PROGRAM main
  VAR
    B1 AT %IX0.0   : BOOL; (* sensor de cajas *)
    KM1 AT %QX0.0  : BOOL; (* banda (bobina 00001 para la PC) *)
    CAJAS AT %MW0  : INT; (* holding 40001: cajas contadas *)
    MARCHA AT %MW1 : INT; (* holding 40002: marcha, la escribe la PC *)
    META AT %MW2   : INT; (* holding 40003: meta de cajas, la escribe la PC *)
    F_CAJA         : R_TRIG;
    CAJA           : BOOL; (* flanco de B1 *)
  END_VAR
  VAR  (* added by the conversion: wires and edge detectors of the diagram *)
    _ADD7_OUT : INT;
    _SEL4_OUT : INT;
    _NE11_OUT : BOOL;
  END_VAR

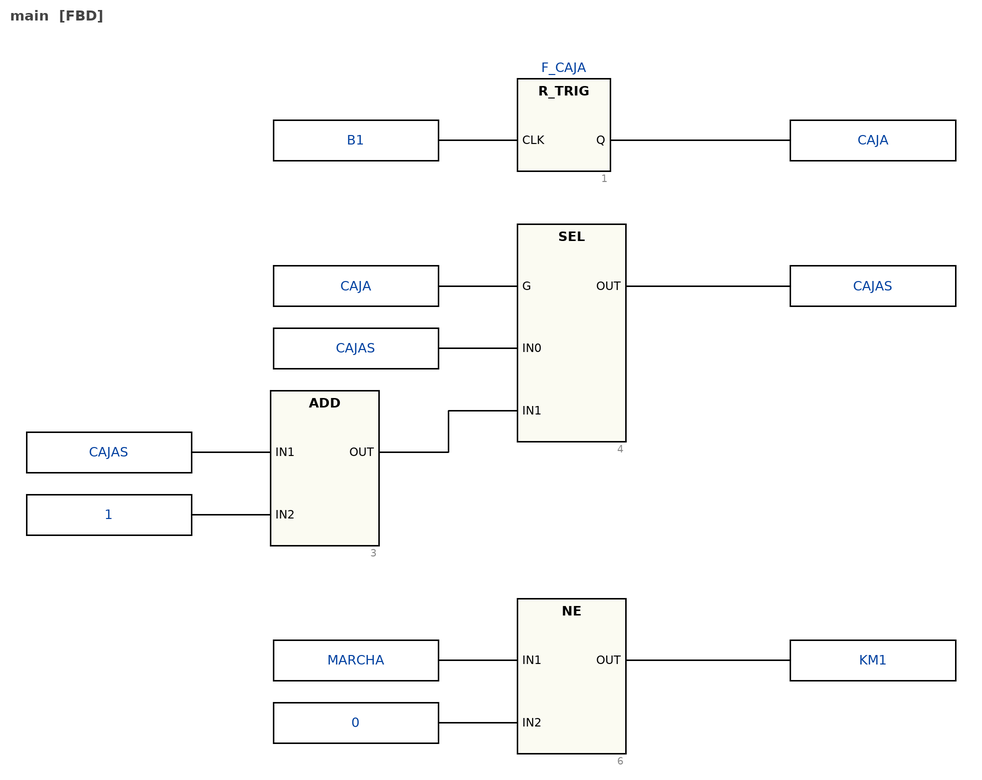
(* FBD diagram, written out as Structured Text *)
F_CAJA(CLK := B1);
CAJA := F_CAJA.Q;
_ADD7_OUT := CAJAS + 1;
_SEL4_OUT := SEL(CAJA, CAJAS, _ADD7_OUT);
CAJAS := _SEL4_OUT;
_NE11_OUT := MARCHA <> 0;
KM1 := _NE11_OUT;
END_PROGRAM
